RoboDK station: Kitting_SSM3_Station.rdk

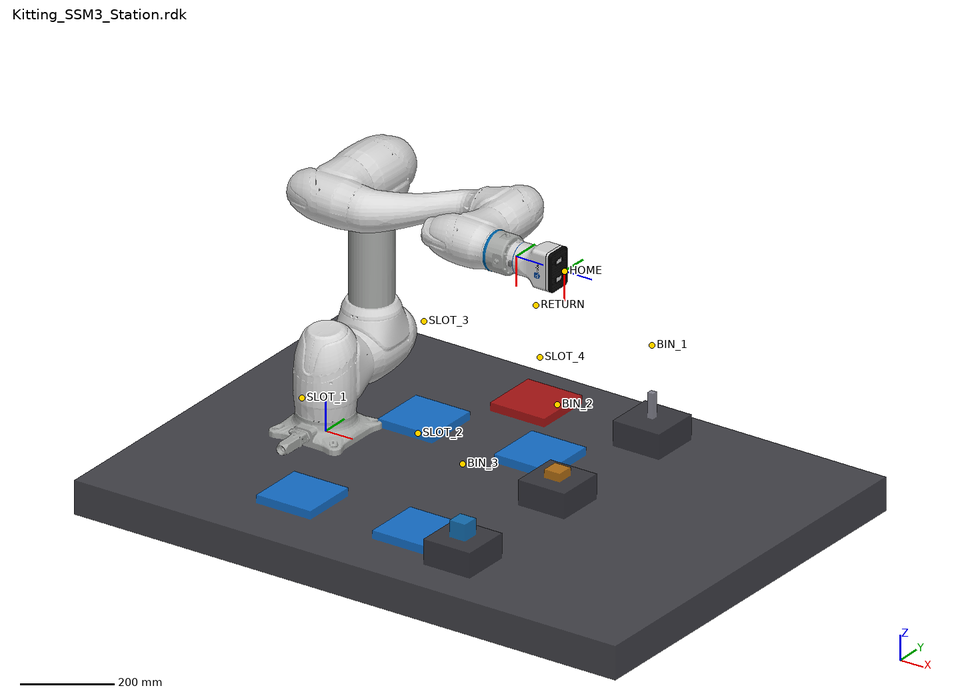
[picture v0: the station drawn from its stored meshes, robots at their saved joint values, targets as dots, program paths as lines]
Station Kitting_SSM3_Station (saved by RoboDK 6.1.1). Poses are relative to the parent item; angles as X-Y-Z fixed-axis rotations.
  - frame Robot_Base at (0, 0, 0) mm
    - robot Doosan Robotics M0609 White: 6 axes, payload 6 kg, reach 900 mm, repeatability 0.03 mm, weight 27 kg
        modified DH rows (alpha deg, a mm, theta deg, d mm): 0, 0, 0, 135; -90, 0, -90, -6.207; 0, 411, -90, 0; -90, 0, 0, 368; 90, 0, 0, 0; -90, 0, 180, 121
        base shift (0, 0, 0) mm, rotated rx 0 ry 0 rz 180 deg
        joint limits [-360, -360, -150, -360, -360, -360] to [360, 360, 150, 360, 360, 360]; home [0, 0, 90, 0, 0, 0]; saved at [0, 0, 90, 0, 0, 0]
      - tool SSM3_Motion_TCP, TCP at (0, 0, 125) mm
      - frame OnRobot-2FG7-Gripper at (0, 0, 0) mm
        - robot OnRobot-2FG7-Gripper-Mechanism: 1 axes
            joint limits [0] to [55]; home [0]; saved at [49.5]
      - frame AUTO_Attach_TCP at (0, 0, 125) mm
  - frame SSM3_Workcell at (0, 0, 0) mm
    - object SSM3_Table at (400, 0, -40) mm, size 1400 x 1000 x 80 mm, geometry from SSM3_Table.stl
    - target HOME (Cartesian target) at (614, 6.21, 546) mm, rotated rx 0 ry 90 rz 0 deg; joints [0, 0, 90, 0, 0, 0] of Doosan Robotics M0609 White
    - object BIN_1_Model at (600, 350, 30) mm, size 120 x 120 x 60 mm, geometry from BIN_1_Model.stl
    - target BIN_1 (Cartesian target) at (600, 350, 230) mm, rotated rx 180 ry 0 rz 0 deg; joints [0, 0, 90, 0, 0, 0] of Doosan Robotics M0609 White
      - object BOLT at (0, 0, 140) mm, rotated rx -180 ry 0 rz 0 deg, size 14 x 14 x 60 mm, geometry from BOLT.stl
    - object BIN_2_Model at (600, 0, 30) mm, size 120 x 120 x 60 mm, geometry from BIN_2_Model.stl
    - target BIN_2 (Cartesian target) at (600, 0, 230) mm, rotated rx 180 ry 0 rz 0 deg; joints [0, 0, 90, 0, 0, 0] of Doosan Robotics M0609 White
      - object SPACER_SHORT at (0, 0, 160) mm, rotated rx -180 ry 0 rz 0 deg, size 40 x 40 x 20 mm, geometry from SPACER_SHORT.stl
    - object BIN_3_Model at (600, -350, 30) mm, size 120 x 120 x 60 mm, geometry from BIN_3_Model.stl
    - target BIN_3 (Cartesian target) at (600, -350, 230) mm, rotated rx 180 ry 0 rz 0 deg; joints [0, 0, 90, 0, 0, 0] of Doosan Robotics M0609 White
      - object SPACER_LONG at (0, 0, 150) mm, rotated rx -180 ry 0 rz 0 deg, size 40 x 40 x 40 mm, geometry from SPACER_LONG.stl
    - object SLOT_1_Model at (150, -300, 10) mm, size 140 x 140 x 20 mm, geometry from SLOT_1_Model.stl
    - target SLOT_1 (Cartesian target) at (150, -300, 240) mm, rotated rx 180 ry 0 rz 0 deg; joints [0, 0, 90, 0, 0, 0] of Doosan Robotics M0609 White
    - object SLOT_2_Model at (450, -300, 10) mm, size 140 x 140 x 20 mm, geometry from SLOT_2_Model.stl
    - target SLOT_2 (Cartesian target) at (450, -300, 240) mm, rotated rx 180 ry 0 rz 0 deg; joints [0, 0, 90, 0, 0, 0] of Doosan Robotics M0609 White
    - object SLOT_3_Model at (150, 150, 10) mm, size 140 x 140 x 20 mm, geometry from SLOT_3_Model.stl
    - target SLOT_3 (Cartesian target) at (150, 150, 240) mm, rotated rx 180 ry 0 rz 0 deg; joints [0, 0, 90, 0, 0, 0] of Doosan Robotics M0609 White
    - object SLOT_4_Model at (450, 150, 10) mm, size 140 x 140 x 20 mm, geometry from SLOT_4_Model.stl
    - target SLOT_4 (Cartesian target) at (450, 150, 240) mm, rotated rx 180 ry 0 rz 0 deg; joints [0, 0, 90, 0, 0, 0] of Doosan Robotics M0609 White
    - object RETURN_Model at (300, 350, 10) mm, size 140 x 140 x 20 mm, geometry from RETURN_Model.stl
    - target RETURN (Cartesian target) at (300, 350, 240) mm, rotated rx 180 ry 0 rz 0 deg; joints [0, 0, 90, 0, 0, 0] of Doosan Robotics M0609 White
